(* IEC 61131-3 sources: codesys-to-astra/src/POUs/F_C2aConcat4, 1 file *)

(* ---- F_C2aConcat4.decl.st ---- *)
// Назначение: замена OSU.CONCAT4 (OwenStringUtils v3.0, с. 39): объединение четырёх строк.
// Автор:      kr0nsch
// Версия:     0.1.0
// Документ:   docs/LIBMAP.md
FUNCTION F_C2aConcat4 : STRING(255)
VAR_INPUT
    sInputString1 : STRING(255);    // строка 1
    sInputString2 : STRING(255);    // строка 2
    sInputString3 : STRING(255);    // строка 3
    sInputString4 : STRING(255);    // строка 4
END_VAR
